    rq_activate_all_grippers(True)
    # end: URCap Program Node
  end
  $ 56 "zero_ftsensor()"
  zero_ftsensor()
  $ 57 "EXTT"
  $ 58 "Set GRP_3F_Enable=Off"
  set_standard_digital_out(4, False)
  $ 59 "Set BarcodeTrigger=Off"
  set_standard_digital_out(6, False)
  $ 60 "Set GRP_3F_Decap=Off"
  set_standard_digital_out(3, False)
  $ 61 "Set GRP_3F_Cap=Off"
  set_standard_digital_out(2, False)
  $ 62 "Set GRP_3F_Open=Off"
  set_standard_digital_out(5, False)
  $ 63 "PSE_T≔get_tool_free_pose(dir=[0,0,0.150], move_in_base_frame=True)"
  global PSE_T=get_tool_free_pose(dir=[0,0,0.150], move_in_base_frame=True)
  $ 64 "If is_reachable(Base_const, [PSE_T])"
  if (is_reachable(p[0.0,0.0,0.0,0.0,0.0,0.0], [PSE_T])):
    $ 65 "MoveL"
    $ 66 "PSE_T" "breakAfter"
    movel(PSE_T, a=1.2, v=0.15)
  end
  while (True):
    $ 67 "Robot Program"
    $ 68 "MAIN"
    $ 69 "command_manager(external_control='uGO', cond_suspend=(ITM_Manipulated and AMR_AtTarget and AMR_Charging and AMR_Battery<40), cond_unsuspend=(AMR_Battery≟60))"
    command_manager(external_control="uGO", cond_suspend=(ITM_Manipulated  and  AMR_AtTarget  and  AMR_Charging  and  AMR_Battery<40), cond_unsuspend=(AMR_Battery == 60))
    $ 70 "log_state(STATE_Info)"
    log_state(STATE_Info)
    $ 71 "Switch STATE"
    switch_1 = STATE
    $ 72 "Case 1"
    if (1 == switch_1):
      $ 73 "Stopping"
      $ 74 "STATE_Info≔'Stopping'"
      global STATE_Info="Stopping"
      $ 75 "end_freedrive_mode()"
      end_freedrive_mode()
      $ 76 "Set"
      set_tcp(p[0.0,0.0,0.161,3.1415,0.0,0.0])
      $ 77 "PSE_T≔get_tool_free_pose(dir=[0,0,0.150], move_in_base_frame=True)"
      global PSE_T=get_tool_free_pose(dir=[0,0,0.150], move_in_base_frame=True)
      $ 78 "If is_reachable(Base_const, [PSE_T])"
      if (is_reachable(p[0.0,0.0,0.0,0.0,0.0,0.0], [PSE_T])):
        $ 79 "MoveL"
        $ 80 "PSE_T" "breakAfter"
        movel(PSE_T, a=1.2, v=0.15)
      end
      $ 81 "do_transition(keep_rxry=OBJ_Picked, r=0)"
      do_transition(keep_rxry=OBJ_Picked, r=0)
      $ 90 "Call Sub_AMR_MiR_V3"
      Sub_AMR_MiR_V3()
      $ 91 "If stopping() and AMR_Done"
      if (stopping()  and  AMR_Done):
        $ 92 "STATE≔2"
        global STATE=2
        $ 93 "ugo_update_outputs()"
        ugo_update_outputs()
      end
    elif (2 == switch_1):
      $ 94 "Case 2"
      $ 95 "Stopped"
      $ 96 "STATE_Info≔'Stopped'"
      global STATE_Info="Stopped"
      $ 97 "Call Sub_AMR_MiR_V3"
      Sub_AMR_MiR_V3()
      $ 98 "If CMD_Reset"
      if (CMD_Reset):
        $ 99 "STATE≔3"
        global STATE=3
        $ 100 "ugo_update_outputs()"
        ugo_update_outputs()
      end
    elif (3 == switch_1):
      $ 101 "Case 3"
      $ 102 " Resetting"
      $ 103 "STATE_Info≔'Resetting'"
      global STATE_Info="Resetting"
      $ 104 "uML"
      $ 105 "reset_error()"
      reset_error()
      $ 106 "reset_warning()"
      reset_warning()
      $ 107 "PROCESS_Step≔0"
      global PROCESS_Step=0
      $ 108 "PROCESS_Info≔''"
      global PROCESS_Info=""
      $ 109 "ARM_Referenced≔ False "
      global ARM_Referenced=  False
      $ 110 "WRK_Done≔ False "
      global WRK_Done=  False
      $ 111 "ITM_Prepared≔ False "
      global ITM_Prepared=  False
      $ 112 "ITM_Manipulated≔ False "
      global ITM_Manipulated=  False
      $ 113 "STP≔0"
      global STP=0
      $ 114 "Action≔0"
      global Action=0
      $ 115 "Action_Info≔''"
      global Action_Info=""
      $ 116 "ITM_ID≔0"
      global ITM_ID=0
      $ 117 "JIG≔0"
      global JIG=0
      $ 118 "JIG_Slot≔0"
      global JIG_Slot=0
      $ 119 "Task_info≔''"
      global Task_info=""
      $ 120 "Set"
      set_tcp(p[0.0,0.0,0.161,3.1415,0.0,0.0])
      $ 121 "App"
      $ 122 "'ADD APPLICATION SPECIFIC COMMANDS'"
      # 'ADD APPLICATION SPECIFIC COMMANDS'
      $ 123 "OBJ_Type≔0"
      global OBJ_Type=0
      $ 124 "OBJ_Nbr≔0"
      global OBJ_Nbr=0
      $ 125 "If CNT_Rack_Output≥50"
      if (CNT_Rack_Output >= 50):
        $ 126 "CNT_Rack_Output≔0"
        global CNT_Rack_Output=0
      end
      $ 127 "TASK≔struct(ID=0, NAVI=struct(target=0, footprint=0, protectiveOff=0, dock=0), WORK=struct(ITM_ID_Src=0, JIG_ID_Src=0, OBJ_Nbr_Src=0, ACT_Src=0, ITM_ID_Tgt=0, JIG_ID_Tgt=0, OBJ_Nbr_Tgt=0, ACT_Tgt=0, OBJ_Type=0))"
      global TASK=struct(ID=0, NAVI=struct(target=0, footprint=0, protectiveOff=0, dock=0), WORK=struct(ITM_ID_Src=0, JIG_ID_Src=0, OBJ_Nbr_Src=0, ACT_Src=0, ITM_ID_Tgt=0, JIG_ID_Tgt=0, OBJ_Nbr_Tgt=0, ACT_Tgt=0, OBJ_Type=0))
      $ 128 "Call Sub_AMR_MiR_V3"
      Sub_AMR_MiR_V3()
      $ 129 "If resetting() and AMR_Done"
      if (resetting()  and  AMR_Done):
        $ 130 "STATE≔4"
        global STATE=4
        $ 131 "ugo_update_outputs()"
        ugo_update_outputs()
      end
    elif (4 == switch_1):
      $ 132 "Case 4"
      $ 133 "Idle"
      $ 134 "STATE_Info≔'Idle'"
      global STATE_Info="Idle"
      $ 135 "If CMD_Start"
      if (CMD_Start):
        $ 136 "STATE≔5"
        global STATE=5
        $ 137 "ugo_update_outputs()"
        ugo_update_outputs()
      end
    elif (5 == switch_1):
      $ 138 "Case 5"
      $ 139 "Starting"
      $ 140 "STATE_Info≔'Starting'"
      global STATE_Info="Starting"
      $ 141 "'ADD COMMANDS WHAT TO START WITH'"
      # 'ADD COMMANDS WHAT TO START WITH'
      $ 142 "Call Sub_AMR_MiR_V3"
      Sub_AMR_MiR_V3()
      $ 143 "get ugo data"
      $ 144 "Assign Tasks"
      $ 145 "TASK.ID = ugo_get_task()"
      TASK.ID = ugo_get_task()
      $ 146 "If TASK.ID≟1"
      if (TASK.ID == 1):
        $ 147 "Task_info≔'Charge'"
        global Task_info="Charge"
        $ 148 "Parameters"
        $ 149 "AMR_PosTarget≔1"
        global AMR_PosTarget=1
      else:
        $ 150 "ElseIf TASK.ID≟9"
        if (TASK.ID == 9):
          $ 151 "'Pick Sarstedt Rack from Variable source'"
          # 'Pick Sarstedt Rack from Variable source'
          $ 152 "Task_info≔'Navigate to Target'"
          global Task_info="Navigate to Target"
          $ 153 "Parameters"
          $ 154 "AMR_PosTarget≔UGO.read_input('00','ITM_ID')"
          global AMR_PosTarget=UGO.read_input("00","ITM_ID")
        else:
          $ 155 "ElseIf TASK.ID≟10"
          if (TASK.ID == 10):
            $ 156 "'Pick Sarstedt Rack from Variable source'"
            # 'Pick Sarstedt Rack from Variable source'
            $ 157 "Task_info≔'Pick Rack'"
            global Task_info="Pick Rack"
            $ 158 "AMR_PosTarget≔2"
            global AMR_PosTarget=2
            $ 159 "Parameters"
            $ 160 "ITM_ID≔UGO.read_input('00','ITM_ID')"
            global ITM_ID=UGO.read_input("00","ITM_ID")
            $ 161 "JIG≔UGO.read_input('00','JIG_ID')"
            global JIG=UGO.read_input("00","JIG_ID")
            $ 162 "OBJ_Type≔3"
            global OBJ_Type=3
          else:
            $ 163 "ElseIf TASK.ID≟11"
            if (TASK.ID == 11):
              $ 164 "'Place Sarstedt Rack on Variable target'"
              # 'Place Sarstedt Rack on Variable target'
              $ 165 "Task_info≔'Place Rack'"
              global Task_info="Place Rack"
              $ 166 "AMR_PosTarget≔2"
              global AMR_PosTarget=2
              $ 167 "Parameters"
              $ 168 "ITM_ID≔UGO.read_input('00','ITM_ID')"
              global ITM_ID=UGO.read_input("00","ITM_ID")
              $ 169 "JIG≔UGO.read_input('00','JIG_ID')"
              global JIG=UGO.read_input("00","JIG_ID")
              $ 170 "OBJ_Type≔3"
              global OBJ_Type=3
            else:
              $ 172 "ElseIf TASK.ID≟12"
              if (TASK.ID == 12):
                $ 173 "Task_info≔'Decapping'"
                global Task_info="Decapping"
                $ 174 "Parameters"
                $ 175 "ITM_ID≔1"
                global ITM_ID=1
                $ 176 "AMR_PosTarget≔AMR_PosActual"
                global AMR_PosTarget=AMR_PosActual
                $ 177 "PRC_TubCounter≔0"
                global PRC_TubCounter=0
              else:
                $ 178 "ElseIf TASK.ID≟13"
                if (TASK.ID == 13):
                  $ 179 "Task_info≔'Empty racks'"
                  global Task_info="Empty racks"
                  $ 180 "Parameters"
                  $ 181 "ITM_ID≔1"
                  global ITM_ID=1
                  $ 182 "AMR_PosTarget≔AMR_PosActual"
                  global AMR_PosTarget=AMR_PosActual
                else:
                  $ 183 "ElseIf TASK.ID≟16"
                  if (TASK.ID == 16):
                    $ 184 "Task_info≔'Decap + Barcode'"
                    global Task_info="Decap + Barcode"
                    $ 185 "Parameters"
                    $ 187 "OBJs_String≔UGO.read_input('00','ObjPos')"
                    global OBJs_String=UGO.read_input("00","ObjPos")
                    $ 188 "OBJs_List≔make_list(length = elements_in_string(OBJs_String), initial_value = -1, capacity = 50)"
                    global OBJs_List=make_list(length = elements_in_string(OBJs_String), initial_value = -1, capacity = 50)
                    $ 189 "OBJs_List≔string_to_list(OBJs_String)"
                    global OBJs_List=string_to_list(OBJs_String)
                    $ 190 "ITM_ID≔1"
                    global ITM_ID=1
                    $ 191 "OBJ_Type≔2"
                    global OBJ_Type=2
                    $ 192 "JIG≔7"
                    global JIG=7
                    $ 193 "AMR_PosTarget≔AMR_PosActual"
                    global AMR_PosTarget=AMR_PosActual
                  else:
                    $ 194 "ElseIf TASK.ID≟30"
                    if (TASK.ID == 30):
                      $ 195 "Task_info≔'Getting bottles'"
                      global Task_info="Getting bottles"
                      $ 196 "Parameters"
                      $ 197 "ITM_ID≔1"
                      global ITM_ID=1
                      $ 198 "OBJ_Type≔4"
                      global OBJ_Type=4
                      $ 199 "JIG≔9"
                      global JIG=9
                      $ 200 "AMR_PosTarget≔4"
                      global AMR_PosTarget=4
                    else:
                      $ 201 "ElseIf TASK.ID≟40"
                      if (TASK.ID == 40):
                        $ 202 "Task_info≔'Placing bottles'"
                        global Task_info="Placing bottles"
                        $ 203 "Parameters"
                        $ 204 "ITM_ID≔1"
                        global ITM_ID=1
                        $ 205 "OBJ_Type≔4"
                        global OBJ_Type=4
                        $ 206 "JIG≔10"
                        global JIG=10
                        $ 207 "AMR_PosTarget≔4"
                        global AMR_PosTarget=4
                      else:
                        $ 208 "ElseIf TASK.ID≟41"
                        if (TASK.ID == 41):
                          $ 209 "Task_info≔'Shaking bottle'"
                          global Task_info="Shaking bottle"
                          $ 210 "Parameters"
                          $ 211 "ITM_ID≔1"
                          global ITM_ID=1
                          $ 212 "OBJ_Type≔4"
                          global OBJ_Type=4
                          $ 213 "JIG≔11"
                          global JIG=11
                          $ 214 "AMR_PosTarget≔4"
                          global AMR_PosTarget=4
                        else:
                          $ 215 "ElseIf TASK.ID≟42"
                          if (TASK.ID == 42):
                            $ 216 "Task_info≔'Decap the bottle'"
                            global Task_info="Decap the bottle"
                            $ 217 "Parameters"
                            $ 218 "ITM_ID≔1"
                            global ITM_ID=1
                            $ 219 "OBJ_Type≔4"
                            global OBJ_Type=4
                            $ 220 "AMR_PosTarget≔4"
                            global AMR_PosTarget=4
                          else:
                            $ 221 "ElseIf TASK.ID≟43"
                            if (TASK.ID == 43):
                              $ 222 "Task_info≔'Pick the Rack'"
                              global Task_info="Pick the Rack"
                              $ 223 "AMR_PosTarget≔5"
                              global AMR_PosTarget=5
                              $ 224 "Parameters"
                              $ 225 "ITM_ID≔UGO.read_input('00','ITM_ID')"
                              global ITM_ID=UGO.read_input("00","ITM_ID")
                              $ 226 "JIG≔UGO.read_input('00','JIG_ID')"
                              global JIG=UGO.read_input("00","JIG_ID")
                              $ 227 "OBJ_Type≔3"
                              global OBJ_Type=3
                            else:
                              $ 228 "ElseIf TASK.ID≟45"
                              if (TASK.ID == 45):
                                $ 229 "Task_info≔'pick the Vial'"
                                global Task_info="pick the Vial"
                                $ 230 "Parameters"
                                $ 231 "ITM_ID≔1"
                                global ITM_ID=1
                                $ 232 "OBJ_Type≔4"
                                global OBJ_Type=4
                                $ 233 "JIG≔12"
                                global JIG=12
                                $ 234 "AMR_PosTarget≔5"
                                global AMR_PosTarget=5
                              else:
                                $ 235 "ElseIf TASK.ID≟46"
                                if (TASK.ID == 46):
                                  $ 236 "Task_info≔'Decap the Vial'"
                                  global Task_info="Decap the Vial"
                                  $ 237 "Parameters"
                                  $ 238 "ITM_ID≔1"
                                  global ITM_ID=1
                                  $ 239 "OBJ_Type≔4"
                                  global OBJ_Type=4
                                  $ 240 "JIG≔13"
                                  global JIG=13
                                  $ 241 "AMR_PosTarget≔5"
                                  global AMR_PosTarget=5
                                else:
                                  $ 242 "ElseIf TASK.ID≟47"
                                  if (TASK.ID == 47):
                                    $ 243 "Task_info≔'Liquid Transfer'"
                                    global Task_info="Liquid Transfer"
                                    $ 244 "Parameters"
                                    $ 245 "ITM_ID≔1"
                                    global ITM_ID=1
                                    $ 246 "OBJ_Type≔4"
                                    global OBJ_Type=4
                                    $ 247 "JIG≔14"
                                    global JIG=14
                                    $ 248 "AMR_PosTarget≔3"
                                    global AMR_PosTarget=3
                                  else:
                                    $ 249 "ElseIf TASK.ID≟48"
                                    if (TASK.ID == 48):
                                      $ 250 "Task_info≔'Place_rack'"
                                      global Task_info="Place_rack"
                                      $ 251 "Parameters"
                                      $ 252 "ITM_ID≔1"
                                      global ITM_ID=1
                                      $ 253 "OBJ_Type≔3"
                                      global OBJ_Type=3
                                      $ 254 "JIG≔7"
                                      global JIG=7
                                      $ 255 "AMR_PosTarget≔5"
                                      global AMR_PosTarget=5
                                    else:
                                      $ 256 "ElseIf TASK.ID≟49"
                                      if (TASK.ID == 49):
                                        $ 257 "Task_info≔'Pick Containers'"
                                        global Task_info="Pick Containers"
                                        $ 258 "Parameters"
                                        $ 259 "ITM_ID≔1"
                                        global ITM_ID=1
                                        $ 260 "OBJ_Type≔6"
                                        global OBJ_Type=6
                                        $ 261 "JIG≔15"
                                        global JIG=15
                                        $ 262 "AMR_PosTarget≔3"
                                        global AMR_PosTarget=3
                                      else:
                                        $ 263 "ElseIf TASK.ID≟50"
                                        if (TASK.ID == 50):
                                          $ 264 "Task_info≔'Decap Containers'"
                                          global Task_info="Decap Containers"
                                          $ 265 "Parameters"
                                          $ 266 "ITM_ID≔1"
                                          global ITM_ID=1
                                          $ 267 "OBJ_Type≔6"
                                          global OBJ_Type=6
                                          $ 268 "JIG≔16"
                                          global JIG=16
                                          $ 269 "AMR_PosTarget≔5"
                                          global AMR_PosTarget=5
                                        else:
                                          $ 270 "ElseIf TASK.ID≟51"
                                          if (TASK.ID == 51):
                                            $ 271 "Task_info≔'Detect Spatula and transfer powder'"
                                            global Task_info="Detect Spatula and transfer powder"
                                            $ 272 "Parameters"
                                            $ 273 "ITM_ID≔1"
                                            global ITM_ID=1
                                            $ 274 "OBJ_Type≔8"
                                            global OBJ_Type=8
                                            $ 275 "JIG≔16"
                                            global JIG=16
                                            $ 276 "AMR_PosTarget≔5"
                                            global AMR_PosTarget=5
                                          else:
                                            $ 277 "ElseIf TASK.ID≟99"
                                            if (TASK.ID == 99):
                                              $ 278 "Task_info≔'Decapping and barcode alignment'"
                                              global Task_info="Decapping and barcode alignment"
                                              $ 279 "Parameters"
                                              $ 280 "PRC_TubNumber≔UGO.read_input('00','TubesNb')"
                                              global PRC_TubNumber=UGO.read_input("00","TubesNb")
                                              $ 281 "PRC_TubCounter≔0"
                                              global PRC_TubCounter=0
                                              $ 282 "ITM_ID≔1"
                                              global ITM_ID=1
                                              $ 283 "AMR_PosTarget≔AMR_PosActual"
                                              global AMR_PosTarget=AMR_PosActual
                                            else:
                                              $ 318 "Else" "noBreak"
                                              $ 319 "set_error(ERROR_WRONG_ORDER)"
                                              set_error(ERROR_WRONG_ORDER)
                                            end
                                          end
                                        end
                                      end
                                    end
                                  end
                                end
                              end
                            end
                          end
                        end
                      end
                    end
                  end
                end
              end
            end
          end
        end
      end
      $ 320 "test ugo"
      $ 321 "Wait: 0.2"
      sleep(0.2)
      $ 322 "ugo_update_outputs()"
      ugo_update_outputs()
      $ 323 "If starting() and AMR_Done"
      if (starting()  and  AMR_Done):
        $ 324 "log_message(Task_info, 'New Task: ')"
        log_message(Task_info, "New Task: ")
        $ 325 "log_message(to_str(TASK.ID), 'Task_ID: ')"
        log_message(to_str(TASK.ID), "Task_ID: ")
        $ 326 "do_transition(keep_rxry=OBJ_Picked)"
        do_transition(keep_rxry=OBJ_Picked)
        $ 327 "STATE≔6"
        global STATE=6
        $ 328 "ugo_update_outputs()"
        ugo_update_outputs()
      end
    elif (6 == switch_1):
      $ 329 "Case 6"
      $ 330 "Execute"
      $ 331 "STATE_Info≔'Execute'"
      global STATE_Info="Execute"
      $ 332 "If  not CMD_Hold and not CMD_Suspend"
      global thread_flag_332=0
      thread Thread_if_332():
        $ 333 "Switch PROCESS_Step"
        switch_2 = PROCESS_Step
        $ 334 "Case 0"
        if (0 == switch_2):
          $ 335 "PROCESS_Info≔'process control'"
          global PROCESS_Info="process control"
          $ 336 "log_process(PROCESS_Info)"
          log_process(PROCESS_Info)
          $ 337 "process control"
          $ 338 "If  not AMR_AtTarget"
          if (  not  AMR_AtTarget):
            $ 339 "PROCESS_Step≔1"
            global PROCESS_Step=1
          else:
            $ 340 "ElseIf (( not ITM_Prepared and  not WRK_Done) or (ITM_Prepared and WRK_Done))"
            if (((  not  ITM_Prepared  and    not  WRK_Done)  or  (ITM_Prepared  and  WRK_Done))):
              $ 341 "PROCESS_Step≔2"
              global PROCESS_Step=2
            else:
              $ 342 "ElseIf  not WRK_Done"
              if (  not  WRK_Done):
                $ 343 "PROCESS_Step≔3"
                global PROCESS_Step=3
              else:
                $ 344 "Else" "noBreak"
                $ 345 "task finished"
                $ 346 "PROCESS_Info≔''"
                global PROCESS_Info=""
                $ 347 "STATE≔7"
                global STATE=7
                $ 348 "ugo_update_outputs()"
                ugo_update_outputs()
              end
            end
          end
        elif (1 == switch_2):
          $ 349 "Case 1"
          $ 350 "navigate"
          $ 351 "'MOVING THE uML'"
          # 'MOVING THE uML'
          $ 352 "PROCESS_Info≔'move to target'"
          global PROCESS_Info="move to target"
          $ 353 "log_process(PROCESS_Info)"
          log_process(PROCESS_Info)
          $ 354 "If TASK.ID≟1"
          if (TASK.ID == 1):
            $ 355 "Action≔51"
            global Action=51
          else:
            $ 356 "Else" "noBreak"
            $ 357 "Action≔52"
            global Action=52
          end
          $ 358 "Call Sub_AMR_MiR_V3"
          Sub_AMR_MiR_V3()
          $ 359 "If AMR_Done"
          if (AMR_Done):
            $ 360 "PROCESS_Step≔0"
            global PROCESS_Step=0
          end
        elif (2 == switch_2):
          $ 361 "Case 2"
          $ 362 "prepare"
          $ 363 "'THINGS THAT HAVE TO BE DONE ONCE IN A SEQUENCE,WORKFLOW'"
          # 'THINGS THAT HAVE TO BE DONE ONCE IN A SEQUENCE,WORKFLOW'
          $ 364 "PROCESS_Info≔'prepare for work'"
          global PROCESS_Info="prepare for work"
          $ 365 "log_process(PROCESS_Info)"
          log_process(PROCESS_Info)
          $ 366 "If TASK.WORK.ITM_ID_Src>1"
          if (TASK.WORK.ITM_ID_Src>1):
            $ 367 "ITM_ID≔TASK.WORK.ITM_ID_Src"
            global ITM_ID=TASK.WORK.ITM_ID_Src
          else:
            $ 368 "ElseIf TASK.WORK.ITM_ID_Tgt>1"
            if (TASK.WORK.ITM_ID_Tgt>1):
              $ 369 "ITM_ID≔TASK.WORK.ITM_ID_Tgt"
              global ITM_ID=TASK.WORK.ITM_ID_Tgt
            end
          end
          $ 370 "If  not ARM_Referenced and (ITM_ID≠0)"
          if (  not  ARM_Referenced  and  (ITM_ID != 0)):
            $ 371 "STP≔1"
            global STP=1
          else:
            $ 372 "ElseIf ARM_Referenced or (ITM_ID≟0)"
            if (ARM_Referenced  or  (ITM_ID == 0)):
              $ 373 "STP≔2"
              global STP=2
            end
          end
          $ 374 "Switch STP"
          switch_3 = STP
          $ 375 "Case 1"
          if (1 == switch_3):
            $ 376 "reference"
            $ 377 "STP_Info≔'reference at target position'"
            global STP_Info="reference at target position"
            $ 378 "log_step(STP_Info)"
            log_step(STP_Info)
            $ 379 "If ITM_ID≟1"
            if (ITM_ID == 1):
              $ 380 "CAM_Done≔ True "
              global CAM_Done=  True
            else:
              $ 381 "Else" "noBreak"
              $ 382 "Action≔131"
              global Action=131
              $ 383 "Call Sub_Vision_V18"
              Sub_Vision_V18()
            end
            $ 385 "If CAM_Done and  not ERROR.FLAG"
            if (CAM_Done  and    not  ERROR.FLAG):
              $ 386 "log_step('ARM referenced')"
              log_step("ARM referenced")
              $ 387 "ARM_Referenced≔ True "
              global ARM_Referenced=  True
            end
          elif (2 == switch_3):
            $ 388 "Case 2"
            $ 389 "manipulate"
            $ 390 "STP_Info≔'manipulate item'"
            global STP_Info="manipulate item"
            $ 391 "log_step(STP_Info)"
            log_step(STP_Info)
            $ 392 "'In case pressing button is needed'"
            # 'In case pressing button is needed'
            $ 393 "If found_in_list(ITM_ID, ITM_ID_List)"
            if (found_in_list(ITM_ID, ITM_ID_List)):
              $ 394 "Switch ITM_ID"
              switch_4 = ITM_ID
              $ 395 "Case 0"
              if (0 == switch_4):
                $ 396 "ITM_Manipulated≔ not ITM_Manipulated"
                global ITM_Manipulated=  not  ITM_Manipulated
              elif (1 == switch_4):
                $ 397 "Case 1"
                $ 398 "ITM_Manipulated≔ not ITM_Manipulated"
                global ITM_Manipulated=  not  ITM_Manipulated
              elif (2 == switch_4):
                $ 399 "Case 2"
              else:
                $ 409 "Default Case"
                $ 410 "ITM_Manipulated≔ not ITM_Manipulated"
                global ITM_Manipulated=  not  ITM_Manipulated
              end
            end
          end
          $ 411 "ITM_Prepared≔(ITM_Manipulated or  not found_in_list(ITM_ID, ITM_ID_List)) and (ARM_Referenced or ITM_ID≟0) and  not WRK_Done"
          global ITM_Prepared=(ITM_Manipulated  or    not  found_in_list(ITM_ID, ITM_ID_List))  and  (ARM_Referenced  or  ITM_ID == 0)  and    not  WRK_Done
          $ 412 "STP≔0"
          global STP=0
          $ 413 "STP_Info≔''"
          global STP_Info=""
          $ 414 "PROCESS_Step≔0"
          global PROCESS_Step=0
        elif (3 == switch_2):
          $ 415 "Case 3"
          $ 416 "work"
          $ 417 "'ADD EVERY MACHINE, OBJECT, STATION TO WORK ON'"
          # 'ADD EVERY MACHINE, OBJECT, STATION TO WORK ON'
          $ 418 "Switch ITM_ID"
          switch_3 = ITM_ID
          $ 419 "Case 1"
          if (1 == switch_3):
            $ 420 "uLM"
            $ 421 "If TASK.ID≟12"
            if (TASK.ID == 12):
              $ 422 "fill racks"
              $ 423 "Action≔151"
              global Action=151
              $ 424 "Call Sub_Vision_V18"
              Sub_Vision_V18()
              $ 425 "If  not ERROR.FLAG"
              if (  not  ERROR.FLAG):
                $ 426 "Actions for the task"
                $ 427 "Action≔1"
                global Action=1
                $ 428 "JIG≔2"
                global JIG=2
                $ 429 "JIG_Slot≔CAM_Result[0]"
                global JIG_Slot=CAM_Result[0]
                $ 430 "OBJ_Nbr≔CAM_Result[0]"
                global OBJ_Nbr=CAM_Result[0]
                $ 431 "OBJ_Type≔2"
                global OBJ_Type=2
                $ 432 "Call Sub_Action_V4"
                Sub_Action_V4()
                $ 433 "If OBJ_Picked"
                if (OBJ_Picked):
                  $ 434 "CAM_Result.remove(0)"
                  CAM_Result.remove(0)
                  $ 435 "PRC_TubCounter≔PRC_TubCounter+1"
                  global PRC_TubCounter=PRC_TubCounter+1
                  $ 436 "If PRC_TubCounter%4≟0"
                  if (PRC_TubCounter%4 == 0):
                    $ 437 "JIG_Slot≔4"
                    global JIG_Slot=4
                  else:
                    $ 438 "Else" "noBreak"
                    $ 439 "JIG_Slot≔PRC_TubCounter%4"
                    global JIG_Slot=PRC_TubCounter%4
                  end
                  $ 440 "OBJ_Nbr≔ceil(PRC_TubCounter/4)"
                  global OBJ_Nbr=ceil(PRC_TubCounter/4)
                  $ 441 "Action≔2"
                  global Action=2
                  $ 442 "JIG≔4"
                  global JIG=4
                  $ 443 "Call Sub_Action_V4"
                  Sub_Action_V4()
                  $ 444 "Action≔151"
                  global Action=151
                  $ 445 "Call Sub_Vision_V18"
                  Sub_Vision_V18()
                end
              end
              $ 446 "If (CAM_Captures≥CAM_PRM_Retries) or (PRC_TubCounter≥32)"
              if ((CAM_Captures >= CAM_PRM_Retries)  or  (PRC_TubCounter >= 32)):
                $ 447 "PROCESS_Step≔0"
                global PROCESS_Step=0
                $ 448 "WRK_Done≔ True "
                global WRK_Done=  True
              end
            else:
              $ 449 "ElseIf TASK.ID≟10"
              if (TASK.ID == 10):
                $ 450 "Pick Rack"
                $ 451 "Action≔131"
                global Action=131
                $ 452 "Call Sub_Vision_V18"
                Sub_Vision_V18()
                $ 453 "Action≔1"
                global Action=1
                $ 454 "Call Sub_Action_V4"
                Sub_Action_V4()
                $ 455 "PROCESS_Step≔0"
                global PROCESS_Step=0
                $ 456 "WRK_Done≔ True "
                global WRK_Done=  True
              else:
                $ 457 "ElseIf TASK.ID≟11"
                if (TASK.ID == 11):
                  $ 458 "Place Rack"
                  $ 459 "Action≔2"
                  global Action=2
                  $ 460 "Call Sub_Action_V4"
                  Sub_Action_V4()
                  $ 461 "PROCESS_Step≔0"
                  global PROCESS_Step=0
                  $ 462 "WRK_Done≔ True "
                  global WRK_Done=  True
                else:
                  $ 463 "ElseIf TASK.ID≟13"
                  if (TASK.ID == 13):
                    $ 464 "empty racks"
                    $ 465 "pick"
                    $ 466 "Action≔1"
                    global Action=1
                    $ 467 "JIG≔4"
                    global JIG=4
                    $ 468 "If PRC_TubCounter%4≟0"
                    if (PRC_TubCounter%4 == 0):
                      $ 469 "JIG_Slot≔4"
                      global JIG_Slot=4
                    else:
                      $ 470 "Else" "noBreak"
                      $ 471 "JIG_Slot≔PRC_TubCounter%4"
                      global JIG_Slot=PRC_TubCounter%4
                    end
                    $ 472 "OBJ_Nbr≔ceil(PRC_TubCounter/4)"
                    global OBJ_Nbr=ceil(PRC_TubCounter/4)
                    $ 473 "OBJ_Type≔2"
                    global OBJ_Type=2
                    $ 474 "Call Sub_Action_V4"
                    Sub_Action_V4()
                    $ 475 "If OBJ_Picked"
                    if (OBJ_Picked):
                      $ 476 "Action≔2"
                      global Action=2
                      $ 477 "JIG≔3"
                      global JIG=3
                      $ 478 "JIG_Slot≔1"
                      global JIG_Slot=1
                      $ 479 "CNT_Rack_Output≔CNT_Rack_Output + 1"
                      global CNT_Rack_Output=CNT_Rack_Output + 1
                      $ 480 "OBJ_Nbr≔CNT_Rack_Output"
                      global OBJ_Nbr=CNT_Rack_Output
                      $ 481 "Call Sub_Action_V4"
                      Sub_Action_V4()
                      $ 482 "If  not ERROR.FLAG"
                      if (  not  ERROR.FLAG):
                        $ 483 "PRC_TubCounter≔PRC_TubCounter - 1"
                        global PRC_TubCounter=PRC_TubCounter - 1
                      end
                    end
                    $ 484 "If CNT_Rack_Output≥50 or PRC_TubCounter≤0"
                    if (CNT_Rack_Output >= 50  or  PRC_TubCounter <= 0):
                      $ 485 "PROCESS_Step≔0"
                      global PROCESS_Step=0
                      $ 486 "WRK_Done≔ True "
                      global WRK_Done=  True
                    end
                  else:
                    $ 487 "ElseIf TASK.ID≟16"
                    if (TASK.ID == 16):
                      $ 488 "CAM_Result≔OBJs_List"
                      global CAM_Result=OBJs_List
                      $ 489 "PRC_CntDetect≔0"
                      global PRC_CntDetect=0
                      $ 490 "Loop PRC_CntDetect<CAM_Result.length()"
                      while (PRC_CntDetect<CAM_Result.length()):
                        $ 491 "Action≔1"
                        global Action=1
                        $ 492 "ITM_ID≔1"
                        global ITM_ID=1
                        $ 493 "JIG≔2"
                        global JIG=2
                        $ 494 "OBJ_Type≔2"
                        global OBJ_Type=2
                        $ 495 "JIG_Slot≔CAM_Result[PRC_CntDetect]"
                        global JIG_Slot=CAM_Result[PRC_CntDetect]
                        $ 496 "OBJ_Nbr≔CAM_Result[PRC_CntDetect]"
                        global OBJ_Nbr=CAM_Result[PRC_CntDetect]
                        $ 497 "Call Sub_Action_V4"
                        Sub_Action_V4()
                        $ 498 "JIG≔1"
                        global JIG=1
                        $ 499 "Action≔11"
                        global Action=11
                        $ 500 "Call Sub_Action_V4"
                        Sub_Action_V4()
                        $ 501 "Action≔12"
                        global Action=12
                        $ 502 "Call Sub_Action_V4"
                        Sub_Action_V4()
                        $ 503 "Action≔6"
                        global Action=6
                        $ 504 "JIG≔6"
                        global JIG=6
                        $ 505 "Call Sub_Action_V4"
                        Sub_Action_V4()
                        $ 506 "Action≔13"
                        global Action=13
                        $ 507 "Call Sub_Action_V4"
                        Sub_Action_V4()
                        $ 508 "Action≔1"
                        global Action=1
                        $ 509 "JIG≔1"
                        global JIG=1
                        $ 510 "Call Sub_Action_V4"
                        Sub_Action_V4()
                        $ 511 "If OBJ_Brc_OK"
                        if (OBJ_Brc_OK):
                          $ 512 "JIG≔2"
                          global JIG=2
                          $ 513 "Action≔2"
                          global Action=2
                          $ 514 "OBJ_Nbr≔CAM_Result[PRC_CntDetect]"
                          global OBJ_Nbr=CAM_Result[PRC_CntDetect]
                          $ 515 "JIG_Slot≔CAM_Result[PRC_CntDetect]"
                          global JIG_Slot=CAM_Result[PRC_CntDetect]
                          $ 516 "OBJ_Type≔2"
                          global OBJ_Type=2
                          $ 517 "Call Sub_Action_V4"
                          Sub_Action_V4()
                        else:
                          $ 518 "Else" "noBreak"
                          $ 519 "Action≔2"
                          global Action=2
                          $ 520 "JIG≔8"
                          global JIG=8
                          $ 521 "Call Sub_Action_V4"
                          Sub_Action_V4()
                        end
                        $ 522 "PRC_CntDetect≔PRC_CntDetect+1"
                        global PRC_CntDetect=PRC_CntDetect+1
                      end
                      $ 523 "PROCESS_Step≔0"
                      global PROCESS_Step=0
                      $ 524 "WRK_Done≔ True "
                      global WRK_Done=  True
                    else:
                      $ 525 "ElseIf TASK.ID≟30"
                      if (TASK.ID == 30):
                        $ 526 "Pick Bottle"
                        $ 527 "Action≔1"
                        global Action=1
                        $ 528 "Call Sub_Action_V4"
                        Sub_Action_V4()
                        $ 529 "PROCESS_Step≔0"
                        global PROCESS_Step=0
                        $ 530 "WRK_Done≔ True "
                        global WRK_Done=  True
                      else:
                        $ 531 "ElseIf TASK.ID≟40"
                        if (TASK.ID == 40):
                          $ 532 "Place Bottle"
                          $ 533 "Action≔2"
                          global Action=2
                          $ 534 "Call Sub_Action_V4"
                          Sub_Action_V4()
                          $ 535 "PROCESS_Step≔0"
                          global PROCESS_Step=0
                          $ 536 "WRK_Done≔ True "
                          global WRK_Done=  True
                        else:
                          $ 537 "ElseIf TASK.ID≟45"
                          if (TASK.ID == 45):
                            $ 538 "Pick Vial"
                            $ 539 "Action≔31"
                            global Action=31
                            $ 540 "Call Sub_Action_V4"
                            Sub_Action_V4()
                            $ 541 "PROCESS_Step≔0"
                            global PROCESS_Step=0
                            $ 542 "WRK_Done≔ True "
                            global WRK_Done=  True
                          else:
                            $ 543 "ElseIf TASK.ID≟46"
                            if (TASK.ID == 46):
                              $ 544 "Decap Vial"
                              $ 545 "Action≔32"
                              global Action=32
                              $ 546 "Call Sub_Action_V4"
                              Sub_Action_V4()
                              $ 547 "PROCESS_Step≔0"
                              global PROCESS_Step=0
                              $ 548 "WRK_Done≔ True "
                              global WRK_Done=  True
                            else:
                              $ 549 "ElseIf TASK.ID≟47"
                              if (TASK.ID == 47):
                                $ 550 "Liquid transfer"
                                $ 551 "Action≔33"
                                global Action=33
                                $ 552 "Call Sub_Action_V4"
                                Sub_Action_V4()
                                $ 553 "PROCESS_Step≔0"
                                global PROCESS_Step=0
                                $ 554 "WRK_Done≔ True "
                                global WRK_Done=  True
                              else:
                                $ 555 "ElseIf TASK.ID≟48"
                                if (TASK.ID == 48):
                                  $ 556 "Place Rack"
                                  $ 557 "Action≔34"
                                  global Action=34
                                  $ 558 "Call Sub_Action_V4"
                                  Sub_Action_V4()
                                  $ 559 "PROCESS_Step≔0"
                                  global PROCESS_Step=0
                                  $ 560 "WRK_Done≔ True "
                                  global WRK_Done=  True
                                else:
                                  $ 561 "ElseIf TASK.ID≟49"
                                  if (TASK.ID == 49):
                                    $ 562 "Pick Powder container"
                                    $ 563 "Action≔35"
                                    global Action=35
                                    $ 564 "Call Sub_Action_V4"
                                    Sub_Action_V4()
                                    $ 565 "PROCESS_Step≔0"
                                    global PROCESS_Step=0
                                    $ 566 "WRK_Done≔ True "
                                    global WRK_Done=  True
                                  else:
                                    $ 567 "ElseIf TASK.ID≟41"
                                    if (TASK.ID == 41):
                                      $ 568 "shake Bottle"
                                      $ 569 "Action≔30"
                                      global Action=30
                                      $ 570 "Call Sub_Action_V4"
                                      Sub_Action_V4()
                                      $ 571 "PROCESS_Step≔0"
                                      global PROCESS_Step=0
                                      $ 572 "WRK_Done≔ True "
                                      global WRK_Done=  True
                                    else:
                                      $ 573 "ElseIf TASK.ID≟42"
                                      if (TASK.ID == 42):
                                        $ 574 "decap the bottle"
                                        $ 575 "Action≔1"
                                        global Action=1
                                        $ 576 "JIG≔9"
                                        global JIG=9
                                        $ 577 "Call Sub_Action_V4"
                                        Sub_Action_V4()
                                        $ 578 "Action≔11"
                                        global Action=11
                                        $ 579 "JIG≔1"
                                        global JIG=1
                                        $ 580 "Call Sub_Action_V4"
                                        Sub_Action_V4()
                                        $ 581 "Action≔12"
                                        global Action=12
                                        $ 582 "JIG≔1"
                                        global JIG=1
                                        $ 583 "Call Sub_Action_V4"
                                        Sub_Action_V4()
                                        $ 584 "Action≔2"
                                        global Action=2
                                        $ 585 "JIG≔8"
                                        global JIG=8
                                        $ 586 "Call Sub_Action_V4"
                                        Sub_Action_V4()
                                        $ 587 "PROCESS_Step≔0"
                                        global PROCESS_Step=0
                                        $ 588 "WRK_Done≔ True "
                                        global WRK_Done=  True
                                      else:
                                        $ 589 "ElseIf TASK.ID≟43"
                                        if (TASK.ID == 43):
                                          $ 590 "Pick the rack"
                                          $ 591 "Action≔131"
                                          global Action=131
                                          $ 592 "Call Sub_Vision_V18"
                                          Sub_Vision_V18()
                                          $ 593 "Action≔1"
                                          global Action=1
                                          $ 594 "Call Sub_Action_V4"
                                          Sub_Action_V4()
                                          $ 595 "PROCESS_Step≔0"
                                          global PROCESS_Step=0
                                          $ 596 "WRK_Done≔ True "
                                          global WRK_Done=  True
                                        else:
                                          $ 597 "ElseIf TASK.ID≟50"
                                          if (TASK.ID == 50):
                                            $ 598 "Decap containers"
                                            $ 599 "Action≔36"
                                            global Action=36
                                            $ 600 "Call Sub_Action_V4"
                                            Sub_Action_V4()
                                            $ 601 "PROCESS_Step≔0"
                                            global PROCESS_Step=0
                                            $ 602 "WRK_Done≔ True "
                                            global WRK_Done=  True
                                          else:
                                            $ 603 "ElseIf TASK.ID≟51"
                                            if (TASK.ID == 51):
                                              $ 604 "Detect Spatula and transfer powder"
                                              $ 605 "Action≔37"
                                              global Action=37
                                              $ 606 "Call Sub_Action_V4"
                                              Sub_Action_V4()
                                              $ 607 "PROCESS_Step≔0"
                                              global PROCESS_Step=0
                                              $ 608 "WRK_Done≔ True "
                                              global WRK_Done=  True
                                            end
                                          end
                                        end
                                      end
                                    end
                                  end
                                end
                              end
                            end
                          end
                        end
                      end
                    end
                  end
                end
              end
            end
          elif (2 == switch_3):
            $ 609 "Case 2"
          elif (5 == switch_3):
            $ 651 "Case 5"
            $ 652 "SarstedtTable"
            $ 653 "Action≔131"
            global Action=131
            $ 654 "Call Sub_Vision_V18"
            Sub_Vision_V18()
            $ 655 "Action≔1"
            global Action=1
            $ 656 "Call Sub_Action_V4"
            Sub_Action_V4()
            $ 657 "PROCESS_Step≔0"
            global PROCESS_Step=0
            $ 658 "WRK_Done≔ True "
            global WRK_Done=  True
          elif (20 == switch_3):
            $ 659 "Case 20"
          elif (43 == switch_3):
            $ 721 "Case 43"
            $ 722 "Pick the rack"
            $ 723 "Action≔131"
            global Action=131
            $ 724 "Call Sub_Vision_V18"
            Sub_Vision_V18()
            $ 725 "Action≔1"
            global Action=1
            $ 726 "Call Sub_Action_V4"
            Sub_Action_V4()
            $ 727 "PROCESS_Step≔0"
            global PROCESS_Step=0
            $ 728 "WRK_Done≔ True "
            global WRK_Done=  True
          else:
            $ 729 "Default Case"
            $ 730 "WRK_Done≔ True "
            global WRK_Done=  True
            $ 731 "PROCESS_Step≔0"
            global PROCESS_Step=0
          end
        end
        thread_flag_332 = 1
      end
      if (  not  CMD_Hold and not CMD_Suspend):
        global thread_handler_332=run Thread_if_332()
        while (thread_flag_332 == 0):
          if not(  not  CMD_Hold and not CMD_Suspend):
            kill thread_handler_332
            thread_flag_332 = 2
          else:
            sync()
          end
        end
      else:
        thread_flag_332 = 2
      end
      $ 732 "If CMD_Hold"
      if (CMD_Hold):
        $ 733 "STATE≔9"
        global STATE=9
        $ 734 "ugo_update_outputs()"
        ugo_update_outputs()
      else:
        $ 735 "ElseIf CMD_Suspend"
        if (CMD_Suspend):
          $ 736 "STATE≔12"
          global STATE=12
          $ 737 "ugo_update_outputs()"
          ugo_update_outputs()
        end
      end
    elif (7 == switch_1):
      $ 738 "Case 7"
      $ 739 "Completing"
      $ 740 "STATE_Info≔'Completing'"
      global STATE_Info="Completing"
      $ 741 "'ADD COMMANDS FOR COMPLETING THE PROCESS'"
      # 'ADD COMMANDS FOR COMPLETING THE PROCESS'
      $ 742 "do_transition(keep_rxry=OBJ_Picked)"
      do_transition(keep_rxry=OBJ_Picked)
      $ 743 "Call Sub_AMR_MiR_V3"
      Sub_AMR_MiR_V3()
      $ 744 "If completing() and AMR_Done"
      if (completing()  and  AMR_Done):
        $ 745 "STATE≔8"
        global STATE=8
        $ 746 "ugo_update_outputs()"
        ugo_update_outputs()
      end
    elif (8 == switch_1):
      $ 747 "Case 8"
      $ 748 "Complete"
      $ 749 "STATE_Info≔'Complete'"
      global STATE_Info="Complete"
      $ 750 "If CMD_Reset"
      if (CMD_Reset):
        $ 751 "STATE≔3"
        global STATE=3
        $ 752 "ugo_update_outputs()"
        ugo_update_outputs()
      end
    elif (9 == switch_1):
      $ 753 "Case 9"
      $ 754 "Holding"
      $ 755 "STATE_Info≔'Holding'"
      global STATE_Info="Holding"
      $ 756 "stopl(0.5)"
      stopl(0.5)
      $ 757 "Call Sub_AMR_MiR_V3"
      Sub_AMR_MiR_V3()
      $ 758 "If holding() and AMR_Done"
      if (holding()  and  AMR_Done):
        $ 759 "STATE≔10"
        global STATE=10
        $ 760 "ugo_update_outputs()"
        ugo_update_outputs()
      end
    elif (10 == switch_1):
      $ 761 "Case 10"
      $ 762 "Held"
      $ 763 "STATE_Info≔'Held'"
      global STATE_Info="Held"
      $ 764 "If CMD_Unhold"
      if (CMD_Unhold):
        $ 765 "end_freedrive_mode()"
        end_freedrive_mode()
        $ 766 "STATE≔11"
        global STATE=11
        $ 767 "ugo_update_outputs()"
        ugo_update_outputs()
      else:
        $ 768 "ElseIf FNC_Freedrive"
        if (FNC_Freedrive):
          $ 769 "freedrive_mode()"
          freedrive_mode()
        else:
          $ 770 "Else" "noBreak"
          $ 771 "end_freedrive_mode()"
          end_freedrive_mode()
        end
      end
    elif (11 == switch_1):
      $ 772 "Case 11"
      $ 773 "Unholding"
      $ 774 "STATE_Info≔'Unholding'"
      global STATE_Info="Unholding"
      $ 775 "Clearing"
      $ 776 "Switch ERROR.ID"
      switch_2 = ERROR.ID
      $ 777 "Case 1002"
      if (1002 == switch_2):
        $ 778 "AMR_AtTarget≔ False "
        global AMR_AtTarget=  False
        $ 779 "ARM_Referenced≔ False "
        global ARM_Referenced=  False
        $ 780 "ITM_Prepared≔ False "
        global ITM_Prepared=  False
        $ 781 "PROCESS_Step≔1"
        global PROCESS_Step=1
      elif (2007 == switch_2):
        $ 782 "Case 2007"
        $ 783 "PROCESS_Step≔1"
        global PROCESS_Step=1
      end
      $ 784 "reset_error()"
      reset_error()
      $ 785 "reset_warning()"
      reset_warning()
      $ 786 "OBJ_Picked≔gripper_has_object()"
      global OBJ_Picked=gripper_has_object()
      $ 787 "Call Sub_AMR_MiR_V3"
      Sub_AMR_MiR_V3()
      $ 788 "If unholding() and AMR_Done"
      if (unholding()  and  AMR_Done):
        $ 789 "STATE≔6"
        global STATE=6
        $ 790 "ugo_update_outputs()"
        ugo_update_outputs()
      end
    elif (12 == switch_1):
      $ 791 "Case 12"
      $ 792 "Suspending"
      $ 793 "STATE_Info≔'Suspending'"
      global STATE_Info="Suspending"
      $ 794 "PROCESS_Info≔str_cat(PROCESS_Info, ' suspended')"
      global PROCESS_Info=str_cat(PROCESS_Info, " suspended")
      $ 795 "If suspending()"
      if (suspending()):
        $ 796 "STATE≔13"
        global STATE=13
        $ 797 "ugo_update_outputs()"
        ugo_update_outputs()
      end
    elif (13 == switch_1):
      $ 798 "Case 13"
      $ 799 "Suspended"
      $ 800 "STATE_Info≔'Suspended'"
      global STATE_Info="Suspended"
      $ 801 "Call Sub_AMR_MiR_V3"
      Sub_AMR_MiR_V3()
      $ 802 "If CMD_Unsuspend"
      if (CMD_Unsuspend):
        $ 803 "STATE≔14"
        global STATE=14
        $ 804 "ugo_update_outputs()"
        ugo_update_outputs()
      end
    elif (14 == switch_1):
      $ 805 "Case 14"
      $ 806 "Unsuspending"
      $ 807 "STATE_Info≔'Unsuspending'"
      global STATE_Info="Unsuspending"
      $ 808 "PROCESS_Step≔0"
      global PROCESS_Step=0
      $ 809 "If unsuspending()"
      if (unsuspending()):
        $ 810 "STATE≔6"
        global STATE=6
        $ 811 "ugo_update_outputs()"
        ugo_update_outputs()
      end
    elif (15 == switch_1):
      $ 812 "Case 15"
      $ 813 "Aborting"
      $ 814 "STATE_Info≔'Aborting'"
      global STATE_Info="Aborting"
      $ 815 "If aborting()"
      if (aborting()):
        $ 816 "STATE≔16"
        global STATE=16
        $ 817 "ugo_update_outputs()"
        ugo_update_outputs()
      end
    elif (16 == switch_1):
      $ 818 "Case 16"
      $ 819 "Aborted"
      $ 820 "STATE_Info≔'Aborted'"
      global STATE_Info="Aborted"
      $ 821 "If CMD_Clear"
      if (CMD_Clear):
        $ 822 "STATE≔17"
        global STATE=17
        $ 823 "ugo_update_outputs()"
        ugo_update_outputs()
      end
    elif (17 == switch_1):
      $ 824 "Case 17"
      $ 825 "Clearing"
      $ 826 "STATE_Info≔'Clearing'"
      global STATE_Info="Clearing"
      $ 827 "Clearing"
      $ 828 "reset_warning()"
      reset_warning()
      $ 829 "reset_error()"
      reset_error()
      $ 830 "If clearing()"
      if (clearing()):
        $ 831 "STATE≔2"
        global STATE=2
        $ 832 "ugo_update_outputs()"
        ugo_update_outputs()
      end
    end
    $ 833 "log_state(STATE_Info)"
    log_state(STATE_Info)
    $ 834 "log_warning(WARNING.MSG)"
    log_warning(WARNING.MSG)
    $ 835 "log_error(ERROR.MSG)"
    log_error(ERROR.MSG)
    $ 836 "Times"
    $ 837 "Switch STATE"
    switch_1 = STATE
    $ 838 "Case 1"
    if (1 == switch_1):
      $ 839 "TM_St_Stopping≔get_time(STATE_Times[STATE-1])"
      global TM_St_Stopping=get_time(STATE_Times[STATE-1])
    elif (2 == switch_1):
      $ 840 "Case 2"
      $ 841 "TM_St_Stopped≔get_time(STATE_Times[STATE-1])"
      global TM_St_Stopped=get_time(STATE_Times[STATE-1])
    elif (3 == switch_1):
      $ 842 "Case 3"
      $ 843 "TM_St_Resetting≔get_time(STATE_Times[STATE-1])"
      global TM_St_Resetting=get_time(STATE_Times[STATE-1])
    elif (4 == switch_1):
      $ 844 "Case 4"
      $ 845 "TM_St_Idle≔get_time(STATE_Times[STATE-1])"
      global TM_St_Idle=get_time(STATE_Times[STATE-1])
    elif (5 == switch_1):
      $ 846 "Case 5"
      $ 847 "TM_St_Starting≔get_time(STATE_Times[STATE-1])"
      global TM_St_Starting=get_time(STATE_Times[STATE-1])
    elif (6 == switch_1):
      $ 848 "Case 6"
      $ 849 "TM_St_Execute≔get_time(STATE_Times[STATE-1])"
      global TM_St_Execute=get_time(STATE_Times[STATE-1])
    elif (7 == switch_1):
      $ 850 "Case 7"
      $ 851 "TM_St_Completin≔get_time(STATE_Times[STATE-1])"
      global TM_St_Completin=get_time(STATE_Times[STATE-1])
    elif (8 == switch_1):
      $ 852 "Case 8"
      $ 853 "TM_St_Complete≔get_time(STATE_Times[STATE-1])"
      global TM_St_Complete=get_time(STATE_Times[STATE-1])
    elif (9 == switch_1):
      $ 854 "Case 9"
      $ 855 "TM_St_Holding≔get_time(STATE_Times[STATE-1])"
      global TM_St_Holding=get_time(STATE_Times[STATE-1])
    elif (10 == switch_1):
      $ 856 "Case 10"
      $ 857 "TM_St_Held≔get_time(STATE_Times[STATE-1])"
      global TM_St_Held=get_time(STATE_Times[STATE-1])
    elif (11 == switch_1):
      $ 858 "Case 11"
      $ 859 "TM_St_Unholding≔get_time(STATE_Times[STATE-1])"
      global TM_St_Unholding=get_time(STATE_Times[STATE-1])
    elif (12 == switch_1):
      $ 860 "Case 12"
      $ 861 "TM_St_Suspendin≔get_time(STATE_Times[STATE-1])"
      global TM_St_Suspendin=get_time(STATE_Times[STATE-1])
    elif (13 == switch_1):
      $ 862 "Case 13"
      $ 863 "TM_St_Suspended≔get_time(STATE_Times[STATE-1])"
      global TM_St_Suspended=get_time(STATE_Times[STATE-1])
    elif (14 == switch_1):
      $ 864 "Case 14"
      $ 865 "TM_St_Unsuspend≔get_time(STATE_Times[STATE-1])"
      global TM_St_Unsuspend=get_time(STATE_Times[STATE-1])
    elif (15 == switch_1):
      $ 866 "Case 15"
      $ 867 "TM_St_Aborting≔get_time(STATE_Times[STATE-1])"
      global TM_St_Aborting=get_time(STATE_Times[STATE-1])
    elif (16 == switch_1):
      $ 868 "Case 16"
      $ 869 "TM_St_Aborted≔get_time(STATE_Times[STATE-1])"
      global TM_St_Aborted=get_time(STATE_Times[STATE-1])
    elif (17 == switch_1):
      $ 870 "Case 17"
      $ 871 "TM_St_Clearing≔get_time(STATE_Times[STATE-1])"
      global TM_St_Clearing=get_time(STATE_Times[STATE-1])
    end
    $ 873 "Wait: 0.1"
    sleep(0.1)
  end
end
